KUKA KRL data list: Main.dat

DEFDAT Main
   ;FOLD EXTERNAL DECLARATIONS;%{PE}%MKUKATPBASIS,%CEXT,%VCOMMON,%P
   ;FOLD BASISTECH EXT;%{PE}%MKUKATPBASIS,%CEXT,%VEXT,%P
   EXT BAS(BAS_COMMAND :IN, REAL :IN)
   DECL INT SUCCESS
   ;ENDFOLD (BASISTECH EXT)
   ;FOLD USER EXT;%{E}%MKUKATPUSER,%CEXT,%VEXT,%P
   ;Make your modifications here

   ;ENDFOLD (USER EXT)
   ;ENDFOLD (EXTERNAL DECLARATIONS)
   DECL PDAT PDEFAULT = { APO_MODE #CDIS, APO_DIST 500.0, VEL 100.0, ACC 35.000, GEAR_JERK 100.0, EXAX_IGN 0 }
   DECL PDAT PPDAT1 = { APO_MODE #CDIS, APO_DIST 500.0, VEL 100.0, ACC 35.000, GEAR_JERK 100.0, EXAX_IGN 0 }
   DECL PDAT PPDAT2 = { APO_MODE #CDIS, APO_DIST 500.0, VEL 100.0, ACC 35.000, GEAR_JERK 100.0, EXAX_IGN 0 }
   DECL PDAT PPDAT3 = { APO_MODE #CDIS, APO_DIST 500.0, VEL 100.0, ACC 35.000, GEAR_JERK 100.0, EXAX_IGN 0 }
   DECL E6POS XUS_A1Turn = { X -108.546845, Y -232.779461, Z 1087.909911, A 64.999963, B 35.0, C 179.999979, S 2, T 34, E1 0.0, E2 0.0, E3 0.0, E4 0.0, E5 0.0, E6 0.0 }
   DECL FDAT FUS_A1Turn = { BASE_NO 0, TOOL_NO 0, IPO_FRAME #BASE, POINT2[] " " }
   DECL E6POS XDS_A1Turn = { X 44.600443, Y -252.941684, Z 1087.909911, A 99.999963, B 35.0, C 179.999979, S 2, T 34, E1 0.0, E2 0.0, E3 0.0, E4 0.0, E5 0.0, E6 0.0 }
   DECL FDAT FDS_A1Turn = { BASE_NO 0, TOOL_NO 0, IPO_FRAME #BASE, POINT2[] " " }
   DECL E6POS XIMM_A1Turn = { X -1.04082929914592E-13, Y 256.843717, Z 1087.909911, A -90.000037, B 35.0, C 179.999979, S 2, T 35, E1 0.0, E2 0.0, E3 0.0, E4 0.0, E5 0.0, E6 0.0 }
   DECL FDAT FIMM_A1Turn = { BASE_NO 0, TOOL_NO 0, IPO_FRAME #BASE, POINT2[] " " }
   DECL LDAT LCPDAT1 = { APO_FAC 50.0, APO_DIST 500.0, AXIS_ACC 35.000, AXIS_VEL 100.0, CIRC_TYP #BASE, JERK_FAC 50.0, ORI_TYP #VAR, VEL 2.0, ACC 35.000, GEAR_JERK 100.0, EXAX_IGN 0 }
   DECL PDAT PPDAT4 = { APO_MODE #CDIS, APO_DIST 500.0, VEL 100.0, ACC 35.000, GEAR_JERK 100.0, EXAX_IGN 0 }
   DECL E6POS XTT_A1Turn = { X 232.779461, Y -108.546845, Z 1087.909911, A 154.999963, B 35.0, C 179.999979, S 2, T 34, E1 0.0, E2 0.0, E3 0.0, E4 0.0, E5 0.0, E6 0.0 }
   DECL FDAT FTT_A1Turn = { BASE_NO 0, TOOL_NO 0, IPO_FRAME #BASE, POINT2[] " " }
   DECL PDAT PPDAT5 = { APO_MODE #CDIS, APO_DIST 500.0, VEL 100.0, ACC 35.000, GEAR_JERK 100.0, EXAX_IGN 0 }
   DECL E6POS XSC_A1Turn = { X 232.779461, Y -108.546845, Z 1087.909911, A 154.999963, B 35.0, C 179.999979, S 2, T 34, E1 0.0, E2 0.0, E3 0.0, E4 0.0, E5 0.0, E6 0.0 }
   DECL FDAT FSC_A1Turn = { BASE_NO 0, TOOL_NO 0, IPO_FRAME #BASE, POINT2[] " " }
ENDDAT
